Staubli VAL3: resfreshPROG.pgx

program resfreshPROG(string x_sHtml)
  local num l_nSize
  local num l_nSize1
  local num l_i
begin
  //call PROGectory:getSize(l_nSize)
  //  call PROGectory:getPROGList(sPROGList)
  call prog:getSize(l_nSize)
  call prog:getProgList(sPROGList)

  if l_nSize>49
    nPgNumPROG=roundUp(l_nSize/49)
  else
    nPgNumPROG=1
  endIf

  l_nSize1=l_nSize%49

  if nPgIndexPROG==nPgNumPROG-1
    if l_nSize1!=0
      resize(sList,1,l_nSize1)
      for l_i = 0 to size(sList)-1
        sList[l_i]=sPROGList[l_i+nPgIndexPROG*49]
      endFor
    else
      resize(sList,1,49)
      for l_i = 0 to size(sList)-1
        sList[l_i]=sPROGList[l_i+nPgIndexPROG*49]
      endFor
    endIf
  else
    resize(sList,1,49)
    for l_i = 0 to size(sList)-1
      sList[l_i]=sPROGList[l_i+nPgIndexPROG*49]
    endFor
  endIf
  userPageBind(x_sHtml,"lst1","options",sList,size(sList),"r")
  sPagePROG=toString("",nPgNumPROG)
  sPgIndexPROG=toString("",nPgIndexPROG+1)
end
